--- copyPoint3.pgx ---
public program copyPoint3(string x_sKey, num x_nTarget, num x_nSource)
  local num l_i
begin
  //2024.12.23 add 增加点位索引
  tTrajBuffer[x_sKey].pPointItem[x_nTarget].pPointRx=trajTemp:tTrajItem[x_sKey].pPointItem[x_nSource].pPointRx
  //tTrajBuffer[x_sKey].pPointItem[x_nTarget].pPointRx[1]=trajTemp:tTrajItem[x_sKey].pPointItem[x_nSource].pPointRx[1]
  tTrajBuffer[x_sKey].pPointItem[x_nTarget].jJointRx=trajTemp:tTrajItem[x_sKey].pPointItem[x_nSource].jJointRx
  tTrajBuffer[x_sKey].pPointItem[x_nTarget].sID=trajTemp:tTrajItem[x_sKey].pPointItem[x_nSource].sID
  tTrajBuffer[x_sKey].pPointItem[x_nTarget].bMarked=trajTemp:tTrajItem[x_sKey].pPointItem[x_nSource].bMarked
  tTrajBuffer[x_sKey].pPointItem[x_nTarget].pInter=trajTemp:tTrajItem[x_sKey].pPointItem[x_nSource].pInter
  tTrajBuffer[x_sKey].pPointItem[x_nTarget].pParaItem.mMdesc=trajTemp:tTrajItem[x_sKey].pPointItem[x_nSource].pParaItem.mMdesc
  tTrajBuffer[x_sKey].pPointItem[x_nTarget].pParaItem.nMoveType=trajTemp:tTrajItem[x_sKey].pPointItem[x_nSource].pParaItem.nMoveType
  tTrajBuffer[x_sKey].pPointItem[x_nTarget].pParaItem.nActionIndex=trajTemp:tTrajItem[x_sKey].pPointItem[x_nSource].pParaItem.nActionIndex
  tTrajBuffer[x_sKey].pPointItem[x_nTarget].pParaItem.nPercentage=trajTemp:tTrajItem[x_sKey].pPointItem[x_nSource].pParaItem.nPercentage
  tTrajBuffer[x_sKey].pPointItem[x_nTarget].pParaItem.nDelay=trajTemp:tTrajItem[x_sKey].pPointItem[x_nSource].pParaItem.nDelay
  tTrajBuffer[x_sKey].pPointItem[x_nTarget].pParaItem.nSigValue=trajTemp:tTrajItem[x_sKey].pPointItem[x_nSource].pParaItem.nSigValue
  tTrajBuffer[x_sKey].pPointItem[x_nTarget].pParaItem.bSafePoint=trajTemp:tTrajItem[x_sKey].pPointItem[x_nSource].pParaItem.bSafePoint
  for l_i = 0 to 2
    tTrajBuffer[x_sKey].pPointItem[x_nTarget].pParaItem.iIfItem.nSigType[l_i]=trajTemp:tTrajItem[x_sKey].pPointItem[x_nSource].pParaItem.iIfItem.nSigType[l_i]
    tTrajBuffer[x_sKey].pPointItem[x_nTarget].pParaItem.iIfItem.nSigIndex[l_i]=trajTemp:tTrajItem[x_sKey].pPointItem[x_nSource].pParaItem.iIfItem.nSigIndex[l_i]
    tTrajBuffer[x_sKey].pPointItem[x_nTarget].pParaItem.iIfItem.nValue[l_i]=trajTemp:tTrajItem[x_sKey].pPointItem[x_nSource].pParaItem.iIfItem.nValue[l_i]
  endFor
  tTrajBuffer[x_sKey].pPointItem[x_nTarget].pParaItem.iIfItem.bANDOR[0]=trajTemp:tTrajItem[x_sKey].pPointItem[x_nSource].pParaItem.iIfItem.bANDOR[0]
  tTrajBuffer[x_sKey].pPointItem[x_nTarget].pParaItem.iIfItem.bANDOR[1]=trajTemp:tTrajItem[x_sKey].pPointItem[x_nSource].pParaItem.iIfItem.bANDOR[1]

end

--- copyPoint31.pgx ---
public program copyPoint31(string x_sKey, num x_nTarget, num x_nSource)
  local num l_i
begin
  //2024.12.23 add 增加点位索引
  trajTemp:tTrajItem[x_sKey].pPointItem[x_nSource].pPointRx=tTrajBuffer[x_sKey].pPointItem[x_nTarget].pPointRx
  trajTemp:tTrajItem[x_sKey].pPointItem[x_nSource].pPointRx[1]=tTrajBuffer[x_sKey].pPointItem[x_nTarget].pPointRx[1]
  trajTemp:tTrajItem[x_sKey].pPointItem[x_nSource].jJointRx=tTrajBuffer[x_sKey].pPointItem[x_nTarget].jJointRx
  trajTemp:tTrajItem[x_sKey].pPointItem[x_nSource].sID=tTrajBuffer[x_sKey].pPointItem[x_nTarget].sID
  trajTemp:tTrajItem[x_sKey].pPointItem[x_nSource].bMarked=tTrajBuffer[x_sKey].pPointItem[x_nTarget].bMarked
  trajTemp:tTrajItem[x_sKey].pPointItem[x_nSource].pInter=tTrajBuffer[x_sKey].pPointItem[x_nTarget].pInter
  trajTemp:tTrajItem[x_sKey].pPointItem[x_nSource].pParaItem.mMdesc=tTrajBuffer[x_sKey].pPointItem[x_nTarget].pParaItem.mMdesc
  trajTemp:tTrajItem[x_sKey].pPointItem[x_nSource].pParaItem.nMoveType=tTrajBuffer[x_sKey].pPointItem[x_nTarget].pParaItem.nMoveType
  trajTemp:tTrajItem[x_sKey].pPointItem[x_nSource].pParaItem.nActionIndex=tTrajBuffer[x_sKey].pPointItem[x_nTarget].pParaItem.nActionIndex
  trajTemp:tTrajItem[x_sKey].pPointItem[x_nSource].pParaItem.nPercentage=tTrajBuffer[x_sKey].pPointItem[x_nTarget].pParaItem.nPercentage
  trajTemp:tTrajItem[x_sKey].pPointItem[x_nSource].pParaItem.nDelay=tTrajBuffer[x_sKey].pPointItem[x_nTarget].pParaItem.nDelay
  trajTemp:tTrajItem[x_sKey].pPointItem[x_nSource].pParaItem.nSigValue=tTrajBuffer[x_sKey].pPointItem[x_nTarget].pParaItem.nSigValue
  trajTemp:tTrajItem[x_sKey].pPointItem[x_nSource].pParaItem.bSafePoint=tTrajBuffer[x_sKey].pPointItem[x_nTarget].pParaItem.bSafePoint
  for l_i = 0 to 2
    trajTemp:tTrajItem[x_sKey].pPointItem[x_nSource].pParaItem.iIfItem.nSigType[l_i]=tTrajBuffer[x_sKey].pPointItem[x_nTarget].pParaItem.iIfItem.nSigType[l_i]
    trajTemp:tTrajItem[x_sKey].pPointItem[x_nSource].pParaItem.iIfItem.nSigIndex[l_i]=tTrajBuffer[x_sKey].pPointItem[x_nTarget].pParaItem.iIfItem.nSigIndex[l_i]
    trajTemp:tTrajItem[x_sKey].pPointItem[x_nSource].pParaItem.iIfItem.nValue[l_i]=tTrajBuffer[x_sKey].pPointItem[x_nTarget].pParaItem.iIfItem.nValue[l_i]
  endFor
  trajTemp:tTrajItem[x_sKey].pPointItem[x_nSource].pParaItem.iIfItem.bANDOR[0]=tTrajBuffer[x_sKey].pPointItem[x_nTarget].pParaItem.iIfItem.bANDOR[0]
  trajTemp:tTrajItem[x_sKey].pPointItem[x_nSource].pParaItem.iIfItem.bANDOR[1]=tTrajBuffer[x_sKey].pPointItem[x_nTarget].pParaItem.iIfItem.bANDOR[1]

end

--- getSize.pgx ---
public program getSize(num& x_nSize)
begin
  // give back the size to trajectory field
  x_nSize=size(trajTemp:tTrajItem)
end

--- getTrajList.pgx ---
public program getTrajList(string& x_sItem[], num x_nIndex)
  local trsf l_tTrsf
  local string l_sItem[6]
  local string l_sEvent
  local string l_sItem2[7]
  local string l_sKey
  local num i
begin
  //  //获取列表
  //  resize(x_sItem,1,1)
  //  l_sKey=first(pt:tCommonStruct)
  //  i=0
  //  while l_sKey!=""
  //    if i!=0
  //      insert(x_sItem[i])
  //    endIf
  //    x_sItem[i]=l_sKey
  //    l_sKey=next(pt:tCommonStruct[l_sKey])
  //    i=i+1
  //    delay(0)
  //  endWhile
  //  if l_sKey=="" and i==0
  //    x_sItem[i]=""
  //  endIf

  //获取列表
  resize(x_sItem,1,x_nIndex)
  l_sKey=first(trajTemp:tTrajItem)
  i=0
  while l_sKey!=""
    x_sItem[i]=l_sKey
    l_sKey=next(trajTemp:tTrajItem[l_sKey])
    i=i+1
  endWhile
  if l_sKey=="" and i==0
    x_sItem[i]=""
  endIf
end

--- stop.pgx ---
program stop()
begin
end
